FUNCTION_BLOCK ControlPanelIn (* Composite Function Block Type *)
  (* Standard: 61499-2 *)
  (* Version 0.0, 7/2/2026, template *)
  PACKAGE Main;
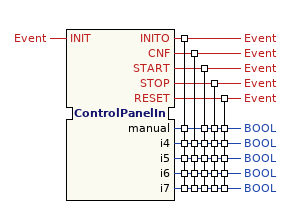
  EVENT_INPUT
    INIT; (* Initialization Request *)
  END_EVENT
  EVENT_OUTPUT
    INITO WITH manual, i4, i5, i6, i7; (* Initialization Confirm *)
    CNF WITH i4, i5, i6, i7; (* Execution Confirmation *)
    START WITH manual, i4, i5, i6, i7;
    STOP WITH manual, i4, i5, i6, i7;
    RESET WITH manual, i4, i5, i6, i7;
  END_EVENT
  VAR_OUTPUT
    manual : BOOL; (* Output event qualifier *)
    i4 : BOOL;
    i5 : BOOL;
    i6 : BOOL;
    i7 : BOOL;
  END_VAR
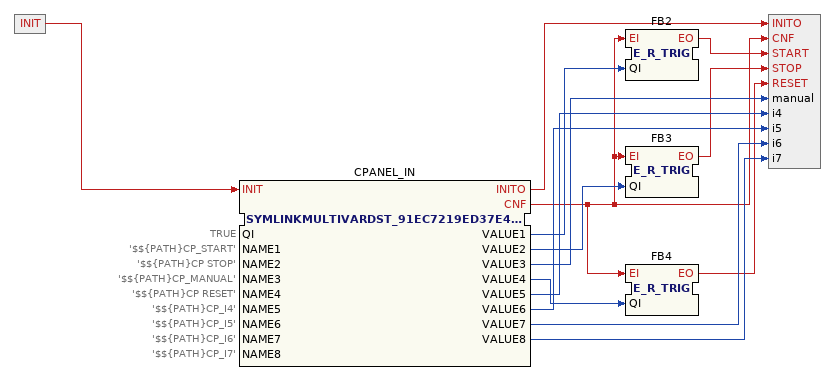
  FBS
    CPANEL_IN : SYMLINKMULTIVARDST_91EC7219ED37E472(QI := TRUE, NAME1 := '$${PATH}CP_START', NAME2 := '$${PATH}CP STOP', NAME3 := '$${PATH}CP_MANUAL', NAME4 := '$${PATH}CP RESET', NAME5 := '$${PATH}CP_I4', NAME6 := '$${PATH}CP_I5', NAME7 := '$${PATH}CP_I6', NAME8 := '$${PATH}CP_I7'); {SET_ATTRIBUTE(Configuration.GenericFBType.InterfaceParams, Runtime.System#I:=8;VALUE${I$}:BOOL,BOOL,BOOL,BOOL,BOOL,BOOL,BOOL,BOOL)}
    FB2 : E_R_TRIG;
    FB3 : E_R_TRIG;
    FB4 : E_R_TRIG;
  END_FBS
  EVENT_CONNECTIONS
    FB3.EO TO STOP;
    FB4.EO TO RESET;
    FB2.EO TO START;
    INIT TO CPANEL_IN.INIT;
    CPANEL_IN.INITO TO INITO;
    CPANEL_IN.CNF TO FB4.EI;
    CPANEL_IN.CNF TO FB3.EI;
    CPANEL_IN.CNF TO FB2.EI;
    CPANEL_IN.CNF TO CNF;
  END_CONNECTIONS
  DATA_CONNECTIONS
    CPANEL_IN.VALUE1 TO FB2.QI;
    CPANEL_IN.VALUE2 TO FB3.QI;
    CPANEL_IN.VALUE3 TO manual;
    CPANEL_IN.VALUE4 TO FB4.QI;
    CPANEL_IN.VALUE5 TO i4;
    CPANEL_IN.VALUE6 TO i5;
    CPANEL_IN.VALUE7 TO i6;
    CPANEL_IN.VALUE8 TO i7;
  END_CONNECTIONS
END_FUNCTION_BLOCK
